Yaskawa INFORM job: MAINPRO.JBI

/JOB
//NAME MAINPRO
//POS
///NPOS 2,0,0,0,0,0
///TOOL 9
///POSTYPE PULSE
///PULSE
C00000=0,0,0,0,0,0
C00001=0,0,0,0,0,0
//INST
///DATE 2026/10/26 01:19
///COMM Generated using RoboDK
///ATTR SC,RW,RJ
///GROUP1 RB1
NOP
'Program generated by Vertical
'Bot Studio for Motoman ES200D
' on 25/10/2026 12:00:00
'Using nominal kinematics.
'Replace objects Replace objec
'ts
'Using Motoman ES200D Base (ta
'rgets wrt base):
'0.0,0.0,0.0,0.0,0.0,0.0
'Setting Tool 9 (Wood_Holder):
SETE P00095 (1) 0
SETE P00095 (2) 0
SETE P00095 (3) 40000
SETE P00095 (4) 0
SETE P00095 (5) 0
SETE P00095 (6) 0
SETTOOL TL#(9) P00095
MOVJ C00000 VJ=50.00
CALL JOB:TAKEPAR
CALL JOB:APPROAC
CALL JOB:SQUARE
CALL JOB:TRANSIT
CALL JOB:CIRCLE
'show Finish_Part1
'hide Part1
CALL JOB:TRANSIT
CALL JOB:STAR
CALL JOB:RETRACT
CALL JOB:DROPPAR
CALL JOB:TAKEPAR
CALL JOB:APPROAC
CALL JOB:SQUARE
CALL JOB:TRANSIT
CALL JOB:CIRCLE
'show Finish_Part2
'hide Part2
CALL JOB:TRANSIT
CALL JOB:STAR
CALL JOB:RETRACT
CALL JOB:DROPPAR
CALL JOB:TAKEPAR
CALL JOB:APPROAC
CALL JOB:SQUARE
CALL JOB:TRANSIT
CALL JOB:CIRCLE
'show Finish_Part3
'hide Part3
CALL JOB:TRANSIT
CALL JOB:STAR
CALL JOB:RETRACT
CALL JOB:DROPPAR
MOVJ C00001 VJ=50.00
END
